(* Logix 5000 project; controller R400_500_XLS vendor 1 type 14 code 216 rev 31.11; software revision 31.01; part 29 of 32 *)
(* tags used below, declared in another part *)
   Abort1 : DINT;   // Not Used
   Alarm : SINT;   // Wait 3 seconds
   ClearIndex : DINT;
   Condenser : INT;
   CondenserHighFlow_1 : BOOL;   // Enables the condenser high flow valve
   CondenserHighFlow_2 : BOOL;   // Enables the condenser high flow valve
   CondenserLowFlow_1 : BOOL;   // Enables the condenser low flow valve
   CondenserLowFlow_2 : BOOL;   // Enables the condenser low flow valve
   CondenserTran : INT;
   CycleSequence : UDT_CYCLE_SEQUENCE;
   DrnSmp : DINT;
   DRYING : DINT;   // Drying id number
   F1rinse : DINT;   // Not Used
   F2rinse : DINT;   // Not Used
   F3rinse : DINT;   // Not Used
   FC06_ONS : DINT;
   FC06Tran1 : BOOL;   // Condition for the wash treatment to start
   FC07Tran1 : BOOL;   // Condition for the rinse treatment to start
   HeatSmp : DINT;
   iFindCRLFIndex : INT;   // Index Of CRLF in String
   iIndexClearMessageOverflowBuffer : INT;   // Message Overflow Buffer is sPrntArray(200-300)
   M : DINT[5];   // Memory Bits
   MinPressRecord : REAL;
   NeutralizationPhaseRequired : BOOL;
   OneShot : DINT[1];
   ONS_FC07 : SINT;
   print_Footer_template : STRING[7];   // Template for the cycle footer
   printTreatString : STRING[85];   // Treatment String
   rIn_WSH61 : REAL;
   Run : DINT;
   sCRLF : STRING;
   Service : DINT[2];   // Unused Service Mode Memory Bit
   sFll_Zero : STRING[20];
   sMessageToPrint : STRING;   // Message To Print
   sOut_WSH61 : STRING;
   sPrntArray : STRING[300];   // Printer String Array
   sResetPrinter : STRING;   // Clears Printer buffer jplv04f ASCII
   sSpaceCharacter : STRING;   // Space Character
   String : STRING[50];   // String
   SumpHeatingStopped : BOOL;   // Sump heating falling edge
   Tmr : TIMER[107];
   Trt_Drying : SINT;
   Trt_PrWsh : DINT;
   Trt_Rinse : DINT;   // Rinse steps
   Trt_Vapor_Exhaust : BOOL;   // Vapor exhaust fan is on
   Trt_Wsh : DINT;
   WSH56_StartHeating : BOOL;   // Start heating
   WSH56_StartPump : BOOL;   // Start pump signal
   WSH56_StartRecirculation : BOOL;   // Start the recirculation
   WSH_35 : BOOL;   // End of neutralization phase
   WshExcBuffer : UDT_WASH;
   AlarmTrigger : INT;   // Triggers the alarm screen if different of 0
   bCycleOrAbortInProcess : BOOL;
   bNewStringDetected : BOOL;
   DateFormat : SINT;   // 0: M-D-Y 1: D-M-Y 2: Y-M-D
   DateTime : DINT[7];
   ENABLE : BOOL;   // Enable bit
   EnaDisPrinter : BOOL;   // Screen 80 Enable/Disable Printer button
   PmpPres : REAL;
   PressureUnit : BOOL;   // Pressure Unit 0=PSIG 1=BAR
   printAlarm : STRING;
   printAlarmMsg : STRING[50];
   PrintChemCondValue : REAL;
   printEvent : STRING[5];
   PrintFrinseCondValue : REAL;
   PrintIndex : DINT;
   sDate : STRING;   // String current date
   sDateTime : STRING;   // String Date Time
   sNullCharacters : STRING;   // Empty String
   SPV_19 : BOOL;   // Screen 80 Enabled/Disabled Pump pressure monitoring
   sTime : STRING;   // String current time
   SumpTemp : REAL;   // Sump temperature in °C
   tStringCopyDebounce : TIMER;
   udtCSVDataLogBatchReport : UDT_CSVDataLog;
   Unit : Hrdwre;   // Unit Configuration
(* MainProgram, continued *)

ROUTINE WSH_56_TRT_WSH   (* ladder *)
// This module calls the routine to perform Wash treatments
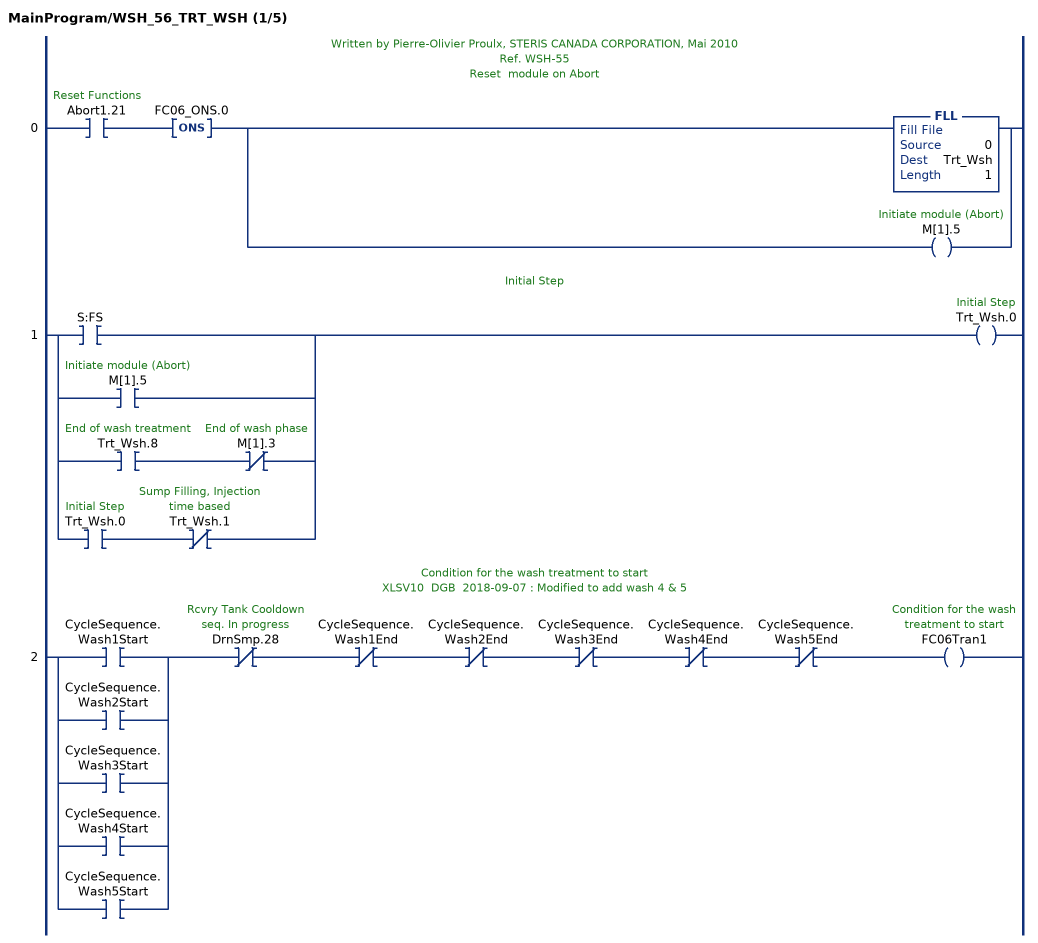
   // Written by Pierre-Olivier Proulx, STERIS CANADA CORPORATION, Mai 2010
   // Ref. WSH-55
   // Reset  module on Abort
   0: XIC(Abort1.21)ONS(FC06_ONS.0)[FLL(0,Trt_Wsh,1) ,OTE(M[1].5) ];
   // Initial Step
   1: [XIC(S:FS) ,XIC(M[1].5) ,XIC(Trt_Wsh.8) XIO(M[1].3) ,XIC(Trt_Wsh.0) XIO(Trt_Wsh.1) ]OTE(Trt_Wsh.0);
   // Condition for the wash treatment to start
   // XLSV10  DGB  2018-09-07 : Modified to add wash 4 & 5
   2: [XIC(CycleSequence.Wash1Start) ,XIC(CycleSequence.Wash2Start) ,XIC(CycleSequence.Wash3Start) ,XIC(CycleSequence.Wash4Start) ,XIC(CycleSequence.Wash5Start) ]XIO(DrnSmp.28)XIO(CycleSequence.Wash1End)XIO(CycleSequence.Wash2End)XIO(CycleSequence.Wash3End)XIO(CycleSequence.Wash4End)XIO(CycleSequence.Wash5End)OTE(FC06Tran1);
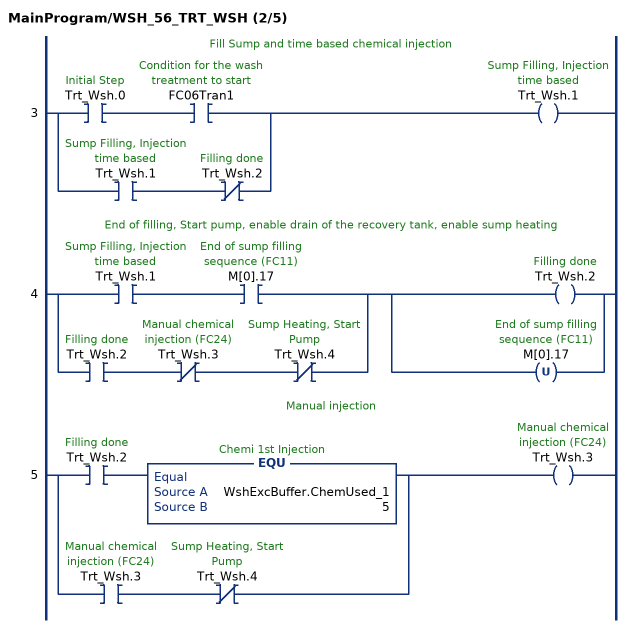
   // Fill Sump and time based chemical injection
   3: [XIC(Trt_Wsh.0) XIC(FC06Tran1) ,XIC(Trt_Wsh.1) XIO(Trt_Wsh.2) ]OTE(Trt_Wsh.1);
   // End of filling, Start pump, enable drain of the recovery tank, enable sump heating
   4: [XIC(Trt_Wsh.1) XIC(M[0].17) ,XIC(Trt_Wsh.2) XIO(Trt_Wsh.3) XIO(Trt_Wsh.4) ][OTE(Trt_Wsh.2) ,OTU(M[0].17) ];
   // Manual injection
   5: [XIC(Trt_Wsh.2) EQU(WshExcBuffer.ChemUsed_1,5) ,XIC(Trt_Wsh.3) XIO(Trt_Wsh.4) ]OTE(Trt_Wsh.3);
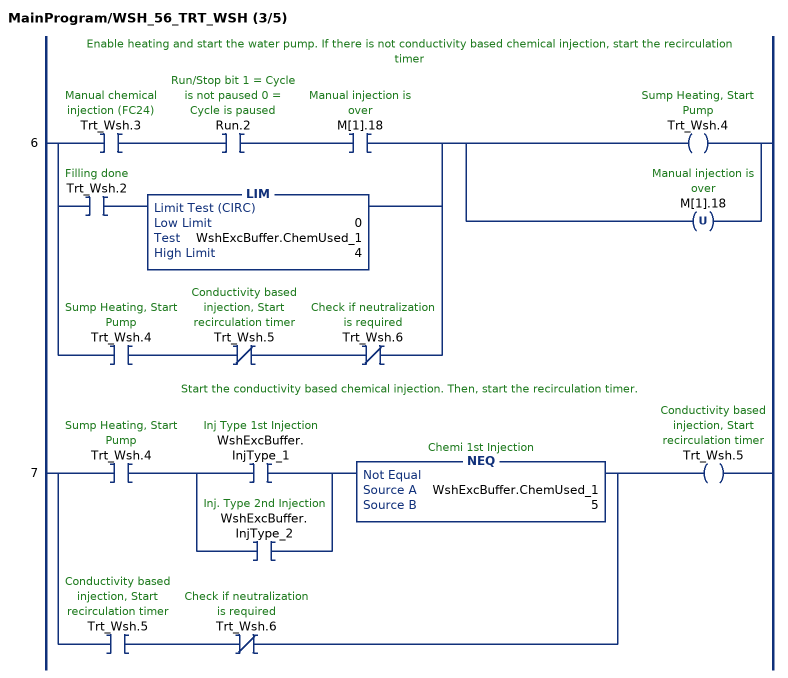
   // Enable heating and start the water pump. If there is not conductivity based chemical injection, start the recirculation timer
   6: [XIC(Trt_Wsh.3) XIC(Run.2) XIC(M[1].18) ,XIC(Trt_Wsh.2) LIM(0,WshExcBuffer.ChemUsed_1,4) ,XIC(Trt_Wsh.4) XIO(Trt_Wsh.5) XIO(Trt_Wsh.6) ][OTE(Trt_Wsh.4) ,OTU(M[1].18) ];
   // Start the conductivity based chemical injection. Then, start the recirculation timer.
   7: [XIC(Trt_Wsh.4) [XIC(WshExcBuffer.InjType_1) ,XIC(WshExcBuffer.InjType_2) ] NEQ(WshExcBuffer.ChemUsed_1,5) ,XIC(Trt_Wsh.5) XIO(Trt_Wsh.6) ]OTE(Trt_Wsh.5);
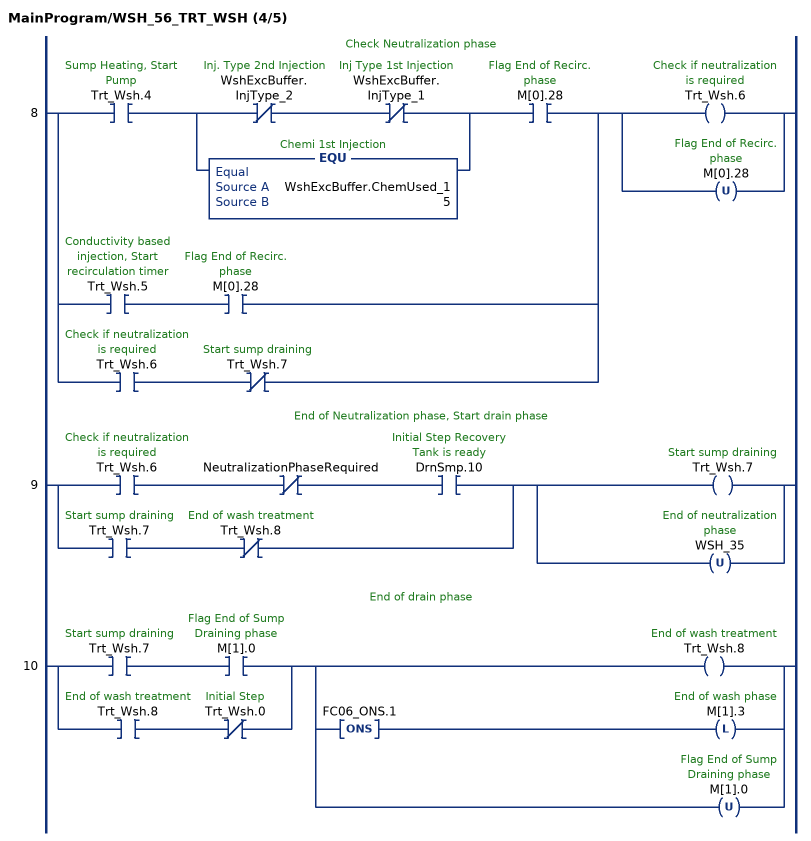
   // Check Neutralization phase
   8: [XIC(Trt_Wsh.4) [XIO(WshExcBuffer.InjType_2) XIO(WshExcBuffer.InjType_1) ,EQU(WshExcBuffer.ChemUsed_1,5) ] XIC(M[0].28) ,XIC(Trt_Wsh.5) XIC(M[0].28) ,XIC(Trt_Wsh.6) XIO(Trt_Wsh.7) ][OTE(Trt_Wsh.6) ,OTU(M[0].28) ];
   // End of Neutralization phase, Start drain phase
   9: [XIC(Trt_Wsh.6) XIO(NeutralizationPhaseRequired) XIC(DrnSmp.10) ,XIC(Trt_Wsh.7) XIO(Trt_Wsh.8) ][OTE(Trt_Wsh.7) ,OTU(WSH_35) ];
   // End of drain phase
   10: [XIC(Trt_Wsh.7) XIC(M[1].0) ,XIC(Trt_Wsh.8) XIO(Trt_Wsh.0) ][OTE(Trt_Wsh.8) ,ONS(FC06_ONS.1) OTL(M[1].3) ,OTU(M[1].0) ];
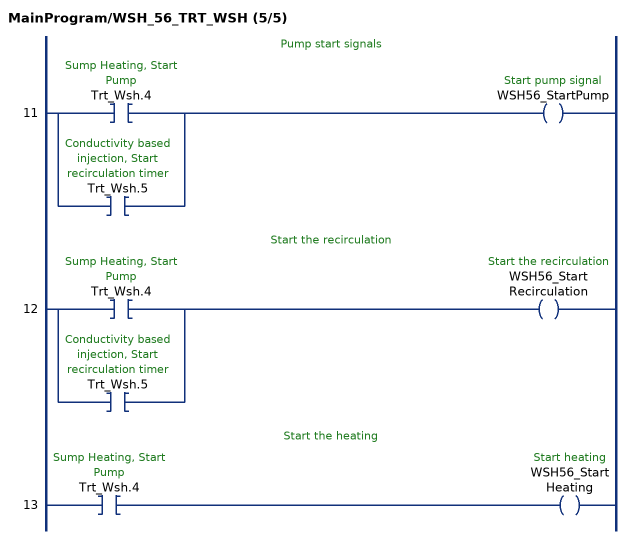
   // Pump start signals
   11: [XIC(Trt_Wsh.4) ,XIC(Trt_Wsh.5) ]OTE(WSH56_StartPump);
   // Start the recirculation
   12: [XIC(Trt_Wsh.4) ,XIC(Trt_Wsh.5) ]OTE(WSH56_StartRecirculation);
   // Start the heating
   13: XIC(Trt_Wsh.4)OTE(WSH56_StartHeating);
END_ROUTINE

ROUTINE WSH_57_TRT_RINSE   (* ladder *)
// This routine performs a rinse treatment.
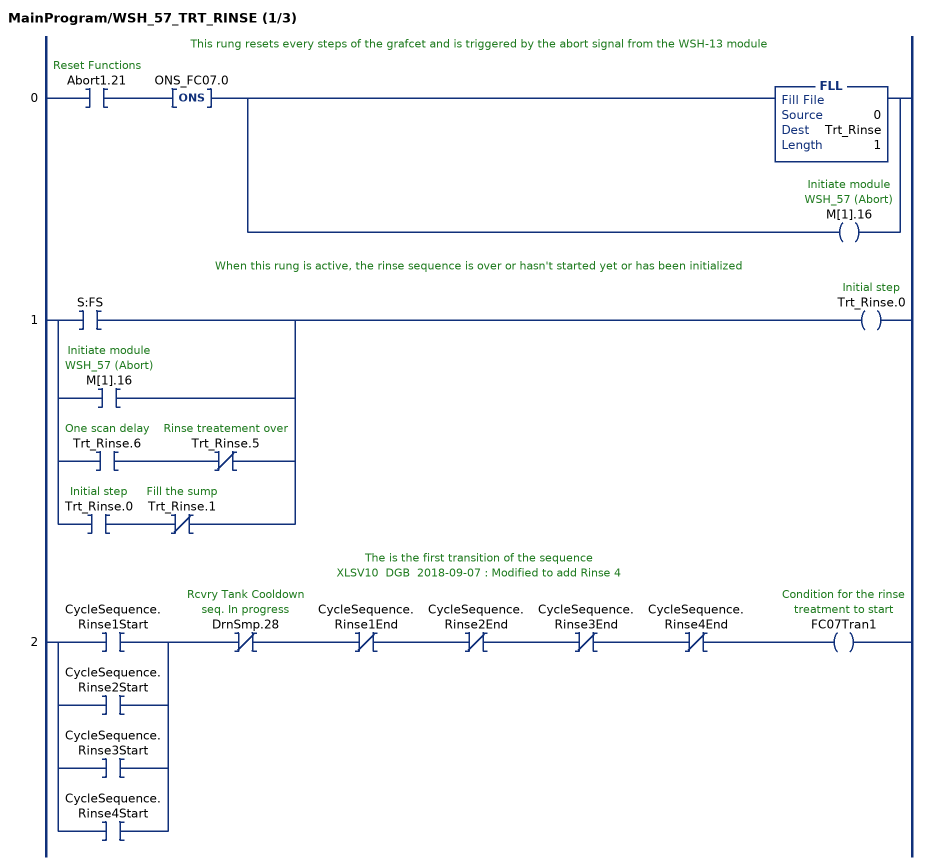
   // This rung resets every steps of the grafcet and is triggered by the abort signal from the WSH-13 module
   0: XIC(Abort1.21)ONS(ONS_FC07.0)[FLL(0,Trt_Rinse,1) ,OTE(M[1].16) ];
   // When this rung is active, the rinse sequence is over or hasn't started yet or has been initialized
   1: [XIC(S:FS) ,XIC(M[1].16) ,XIC(Trt_Rinse.6) XIO(Trt_Rinse.5) ,XIC(Trt_Rinse.0) XIO(Trt_Rinse.1) ]OTE(Trt_Rinse.0);
   // The is the first transition of the sequence
   // XLSV10  DGB  2018-09-07 : Modified to add Rinse 4
   2: [XIC(CycleSequence.Rinse1Start) ,XIC(CycleSequence.Rinse2Start) ,XIC(CycleSequence.Rinse3Start) ,XIC(CycleSequence.Rinse4Start) ]XIO(DrnSmp.28)XIO(CycleSequence.Rinse1End)XIO(CycleSequence.Rinse2End)XIO(CycleSequence.Rinse3End)XIO(CycleSequence.Rinse4End)OTE(FC07Tran1);
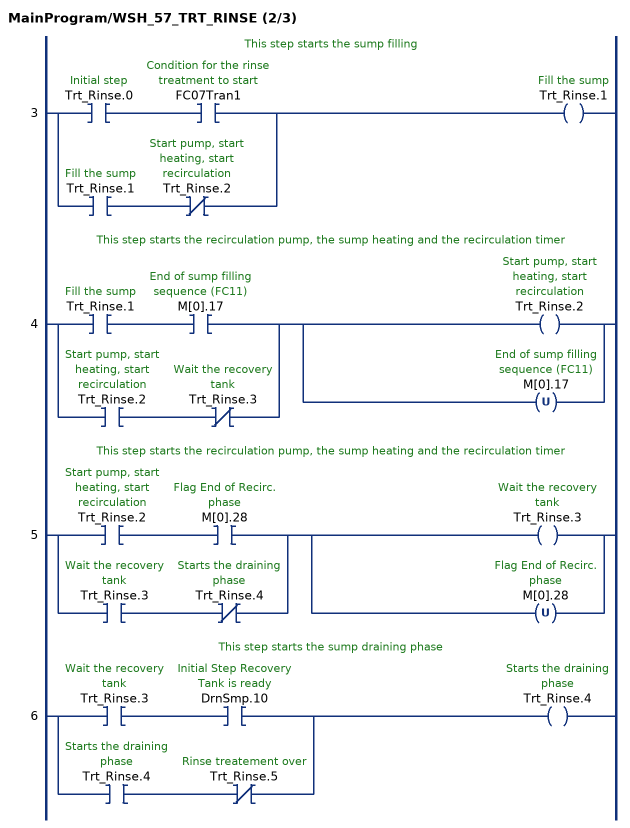
   // This step starts the sump filling
   3: [XIC(Trt_Rinse.0) XIC(FC07Tran1) ,XIC(Trt_Rinse.1) XIO(Trt_Rinse.2) ]OTE(Trt_Rinse.1);
   // This step starts the recirculation pump, the sump heating and the recirculation timer
   4: [XIC(Trt_Rinse.1) XIC(M[0].17) ,XIC(Trt_Rinse.2) XIO(Trt_Rinse.3) ][OTE(Trt_Rinse.2) ,OTU(M[0].17) ];
   // This step starts the recirculation pump, the sump heating and the recirculation timer
   5: [XIC(Trt_Rinse.2) XIC(M[0].28) ,XIC(Trt_Rinse.3) XIO(Trt_Rinse.4) ][OTE(Trt_Rinse.3) ,OTU(M[0].28) ];
   // This step starts the sump draining phase
   6: [XIC(Trt_Rinse.3) XIC(DrnSmp.10) ,XIC(Trt_Rinse.4) XIO(Trt_Rinse.5) ]OTE(Trt_Rinse.4);
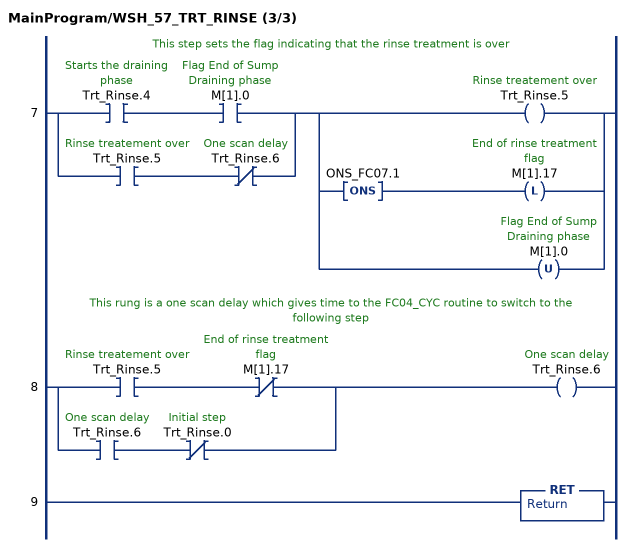
   // This step sets the flag indicating that the rinse treatment is over
   7: [XIC(Trt_Rinse.4) XIC(M[1].0) ,XIC(Trt_Rinse.5) XIO(Trt_Rinse.6) ][OTE(Trt_Rinse.5) ,ONS(ONS_FC07.1) OTL(M[1].17) ,OTU(M[1].0) ];
   // This rung is a one scan delay which gives time to the FC04_CYC routine to switch to the following step
   8: [XIC(Trt_Rinse.5) XIO(M[1].17) ,XIC(Trt_Rinse.6) XIO(Trt_Rinse.0) ]OTE(Trt_Rinse.6);
   9: RET();
END_ROUTINE

ROUTINE WSH_59_CONDENSER_WET   (* ladder *)
// This routine manages the condenser operation
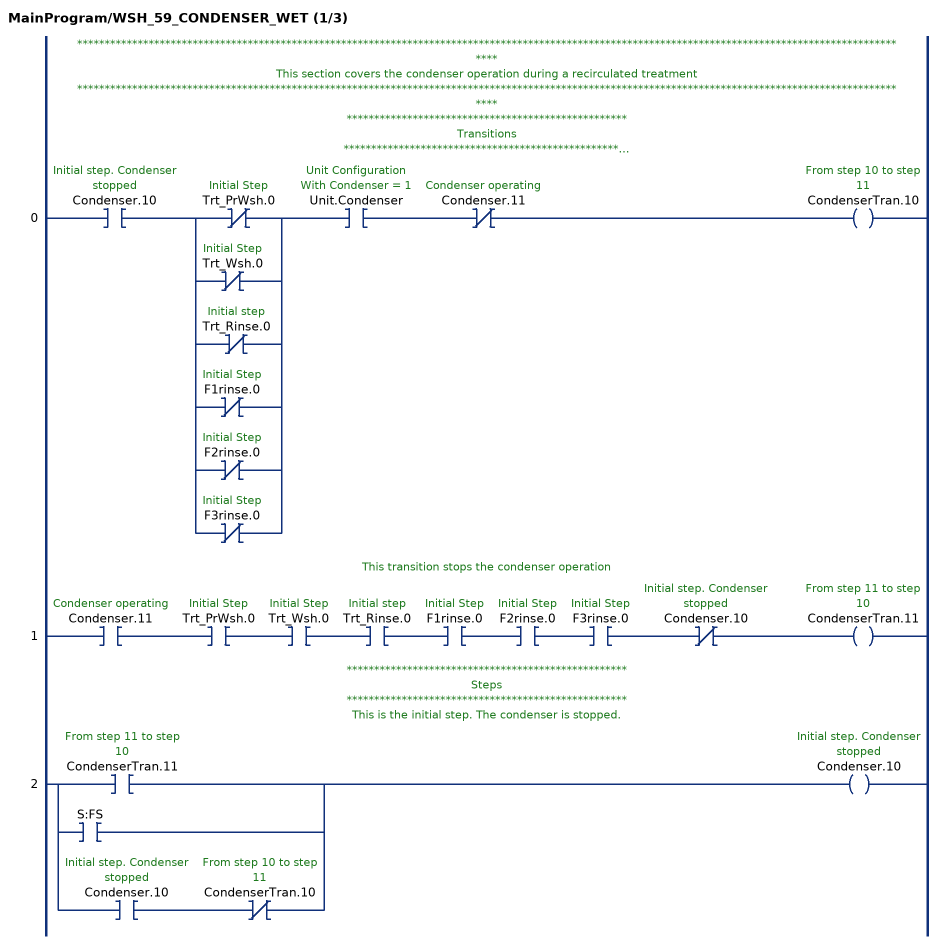
   // *********************************************************************************************************************************************************
   // This section covers the condenser operation during a recirculated treatment
   // *********************************************************************************************************************************************************
   // ***************************************************
   // Transitions
   // ***************************************************
   // This condition triggers the condenser operation
   0: XIC(Condenser.10)[XIO(Trt_PrWsh.0) ,XIO(Trt_Wsh.0) ,XIO(Trt_Rinse.0) ,XIO(F1rinse.0) ,XIO(F2rinse.0) ,XIO(F3rinse.0) ]XIC(Unit.Condenser)XIO(Condenser.11)OTE(CondenserTran.10);
   // This transition stops the condenser operation
   1: XIC(Condenser.11)XIC(Trt_PrWsh.0)XIC(Trt_Wsh.0)XIC(Trt_Rinse.0)XIC(F1rinse.0)XIC(F2rinse.0)XIC(F3rinse.0)XIO(Condenser.10)OTE(CondenserTran.11);
   // ***************************************************
   // Steps
   // ***************************************************
   // This is the initial step. The condenser is stopped.
   2: [XIC(CondenserTran.11) ,XIC(S:FS) ,XIC(Condenser.10) XIO(CondenserTran.10) ]OTE(Condenser.10);
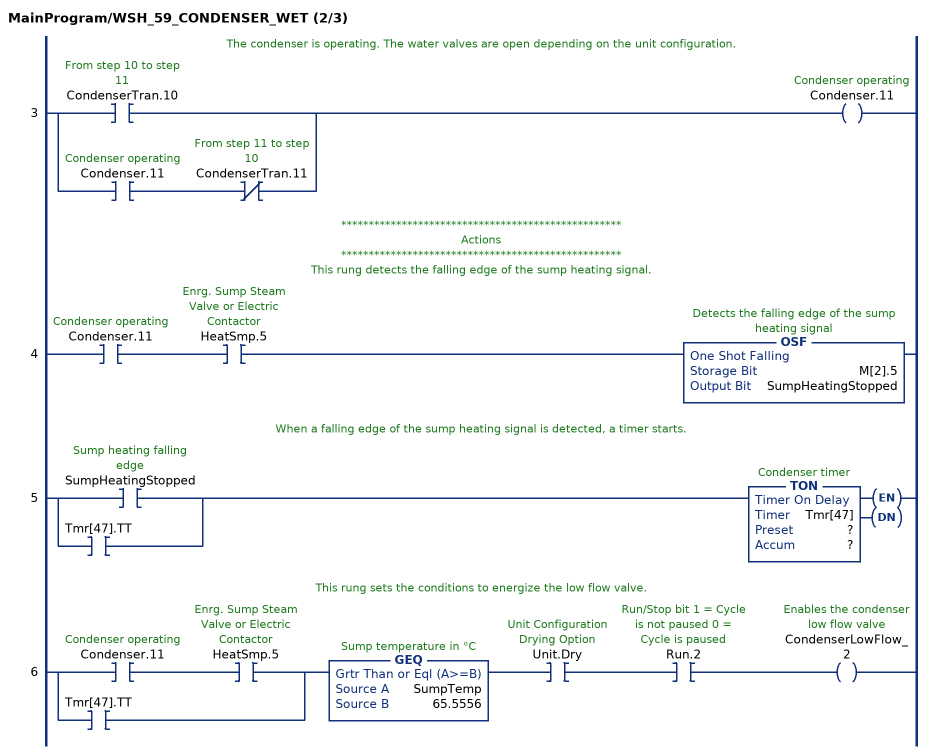
   // The condenser is operating. The water valves are open depending on the unit configuration.
   3: [XIC(CondenserTran.10) ,XIC(Condenser.11) XIO(CondenserTran.11) ]OTE(Condenser.11);
   // ***************************************************
   // Actions
   // ***************************************************
   // This rung detects the falling edge of the sump heating signal.
   4: XIC(Condenser.11)XIC(HeatSmp.5)OSF(M[2].5,SumpHeatingStopped);
   // When a falling edge of the sump heating signal is detected, a timer starts.
   5: [XIC(SumpHeatingStopped) ,XIC(Tmr[47].TT) ]TON(Tmr[47],?,?);
   // This rung sets the conditions to energize the low flow valve.
   6: [XIC(Condenser.11) XIC(HeatSmp.5) ,XIC(Tmr[47].TT) ]GEQ(SumpTemp,65.5556)XIC(Unit.Dry)XIC(Run.2)OTE(CondenserLowFlow_2);
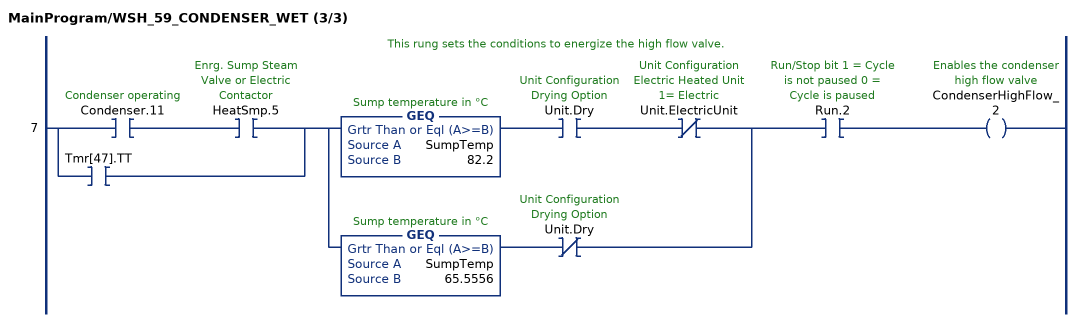
   // This rung sets the conditions to energize the high flow valve.
   7: [XIC(Condenser.11) XIC(HeatSmp.5) ,XIC(Tmr[47].TT) ][GEQ(SumpTemp,82.2) XIC(Unit.Dry) XIO(Unit.ElectricUnit) ,GEQ(SumpTemp,65.5556) XIO(Unit.Dry) ]XIC(Run.2)OTE(CondenserHighFlow_2);
END_ROUTINE

ROUTINE WSH_60_CONDENSER_DRY_VENT   (* ladder *)
// This routine manages the condenser operation
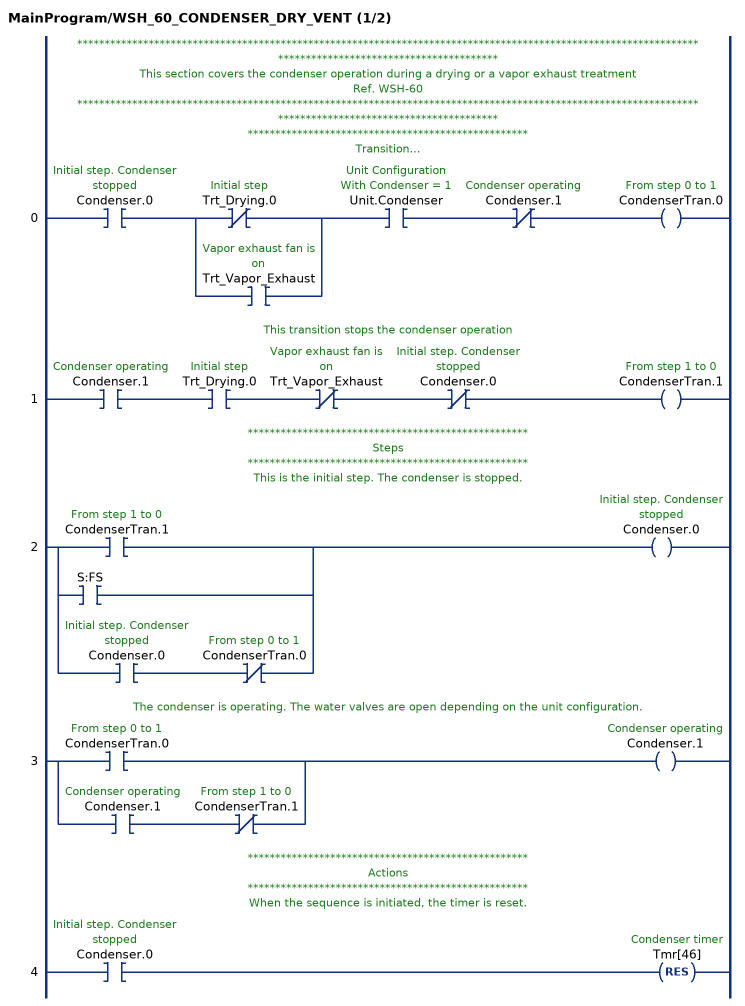
   // *********************************************************************************************************************************************************
   // This section covers the condenser operation during a drying or a vapor exhaust treatment
   // Ref. WSH-60
   // *********************************************************************************************************************************************************
   // ***************************************************
   // Transitions
   // ***************************************************
   // This condition triggers the condenser operation
   0: XIC(Condenser.0)[XIO(Trt_Drying.0) ,XIC(Trt_Vapor_Exhaust) ]XIC(Unit.Condenser)XIO(Condenser.1)OTE(CondenserTran.0);
   // This transition stops the condenser operation
   1: XIC(Condenser.1)XIC(Trt_Drying.0)XIO(Trt_Vapor_Exhaust)XIO(Condenser.0)OTE(CondenserTran.1);
   // ***************************************************
   // Steps
   // ***************************************************
   // This is the initial step. The condenser is stopped.
   2: [XIC(CondenserTran.1) ,XIC(S:FS) ,XIC(Condenser.0) XIO(CondenserTran.0) ]OTE(Condenser.0);
   // The condenser is operating. The water valves are open depending on the unit configuration.
   3: [XIC(CondenserTran.0) ,XIC(Condenser.1) XIO(CondenserTran.1) ]OTE(Condenser.1);
   // ***************************************************
   // Actions
   // ***************************************************
   // When the sequence is initiated, the timer is reset.
   4: XIC(Condenser.0)RES(Tmr[46]);
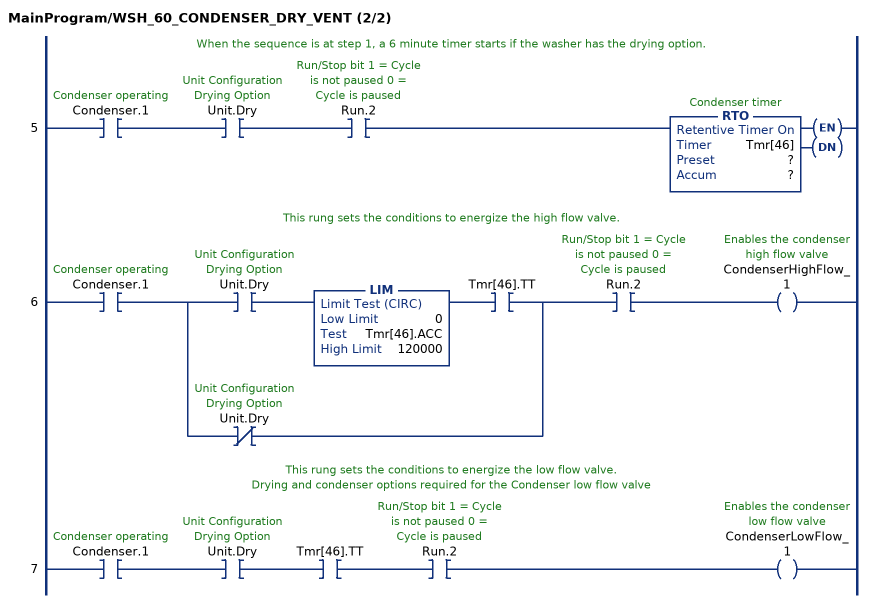
   // When the sequence is at step 1, a 6 minute timer starts if the washer has the drying option.
   5: XIC(Condenser.1)XIC(Unit.Dry)XIC(Run.2)RTO(Tmr[46],?,?);
   // This rung sets the conditions to energize the high flow valve.
   6: XIC(Condenser.1)[XIC(Unit.Dry) LIM(0,Tmr[46].ACC,120000) XIC(Tmr[46].TT) ,XIO(Unit.Dry) ]XIC(Run.2)OTE(CondenserHighFlow_1);
   // This rung sets the conditions to energize the low flow valve.
   // Drying and condenser options required for the Condenser low flow valve
   7: XIC(Condenser.1)XIC(Unit.Dry)XIC(Tmr[46].TT)XIC(Run.2)OTE(CondenserLowFlow_1);
END_ROUTINE

ROUTINE WSH_61_PRINT_STRING_ELEMENT   (* ladder *)
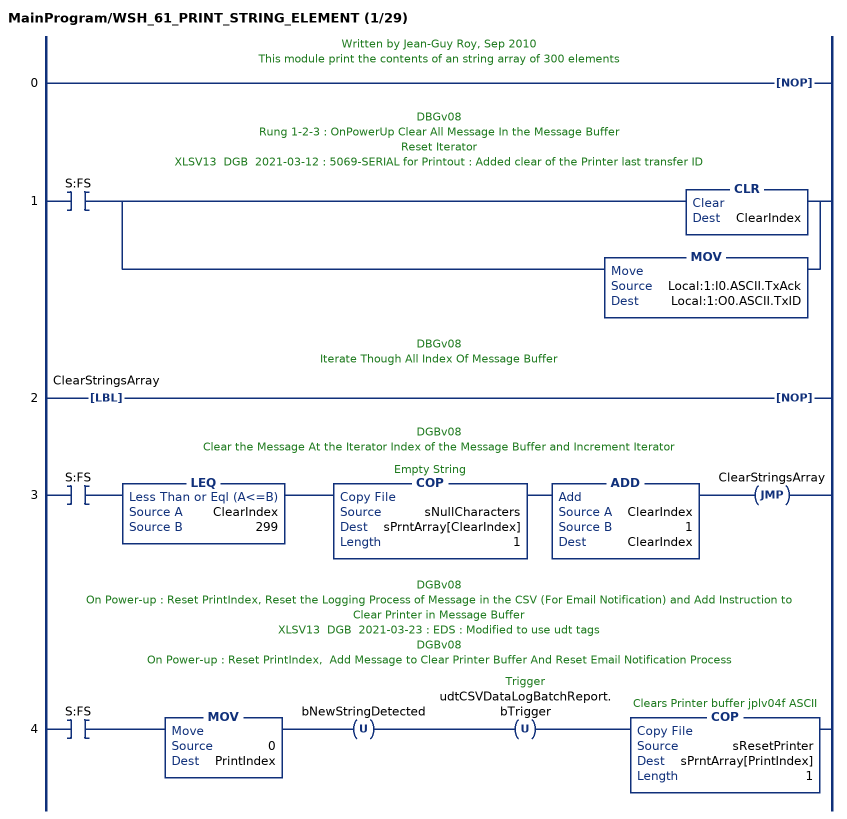
   // Written by Jean-Guy Roy, Sep 2010
   // This module print the contents of an string array of 300 elements
   0: NOP();
   // DBGv08
   // Rung 1-2-3 : OnPowerUp Clear All Message In the Message Buffer
   // Reset Iterator
   // XLSV13  DGB  2021-03-12 : 5069-SERIAL for Printout : Added clear of the Printer last transfer ID
   1: XIC(S:FS)[CLR(ClearIndex) ,MOV(Local:1:I0.ASCII.TxAck,Local:1:O0.ASCII.TxID) ];
   // DBGv08
   // Iterate Though All Index Of Message Buffer
   2: LBL(ClearStringsArray)NOP();
   // DGBv08
   // Clear the Message At the Iterator Index of the Message Buffer and Increment Iterator
   3: XIC(S:FS)LEQ(ClearIndex,299)COP(sNullCharacters,sPrntArray[ClearIndex],1)ADD(ClearIndex,1,ClearIndex)JMP(ClearStringsArray);
   // DGBv08
   // On Power-up : Reset PrintIndex, Reset the Logging Process of Message in the CSV (For Email Notification) and Add Instruction to Clear Printer in Message Buffer
   // XLSV13  DGB  2021-03-23 : EDS : Modified to use udt tags
   // DGBv08
   // On Power-up : Reset PrintIndex,  Add Message to Clear Printer Buffer And Reset Email Notification Process
   4: XIC(S:FS)MOV(0,PrintIndex)OTU(bNewStringDetected)OTU(udtCSVDataLogBatchReport.bTrigger)COP(sResetPrinter,sPrntArray[PrintIndex],1);
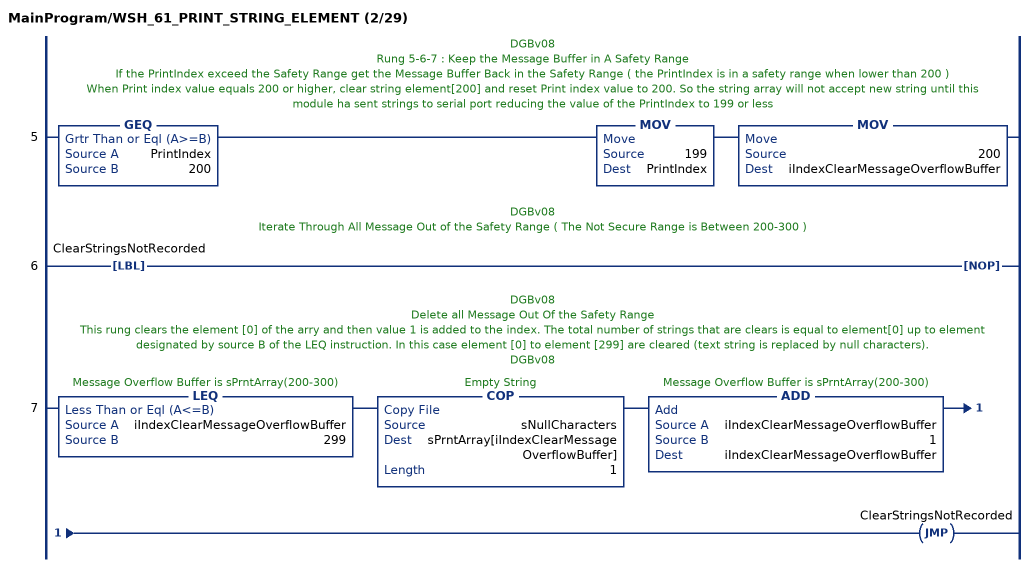
   // DGBv08
   // Rung 5-6-7 : Keep the Message Buffer in A Safety Range
   // If the PrintIndex exceed the Safety Range get the Message Buffer Back in the Safety Range ( the PrintIndex is in a safety range when lower than 200 )
   // When Print index value equals 200 or higher, clear string element[200] and reset Print index value to 200. So the string array will not accept new string until this module ha sent strings to serial port reducing the value of the PrintIndex to 199 or less
   5: GEQ(PrintIndex,200)MOV(199,PrintIndex)MOV(200,iIndexClearMessageOverflowBuffer);
   // DGBv08
   // Iterate Through All Message Out of the Safety Range ( The Not Secure Range is Between 200-300 )
   6: LBL(ClearStringsNotRecorded)NOP();
   // DGBv08
   // Delete all Message Out Of the Safety Range
   // This rung clears the element [0] of the arry and then value 1 is added to the index. The total number of strings that are clears is equal to element[0] up to element designated by source B of the LEQ instruction. In this case element [0] to element [299] are cleared (text string is replaced by null characters).
   // DGBv08
   7: LEQ(iIndexClearMessageOverflowBuffer,299)COP(sNullCharacters,sPrntArray[iIndexClearMessageOverflowBuffer],1)ADD(iIndexClearMessageOverflowBuffer,1,iIndexClearMessageOverflowBuffer)JMP(ClearStringsNotRecorded);
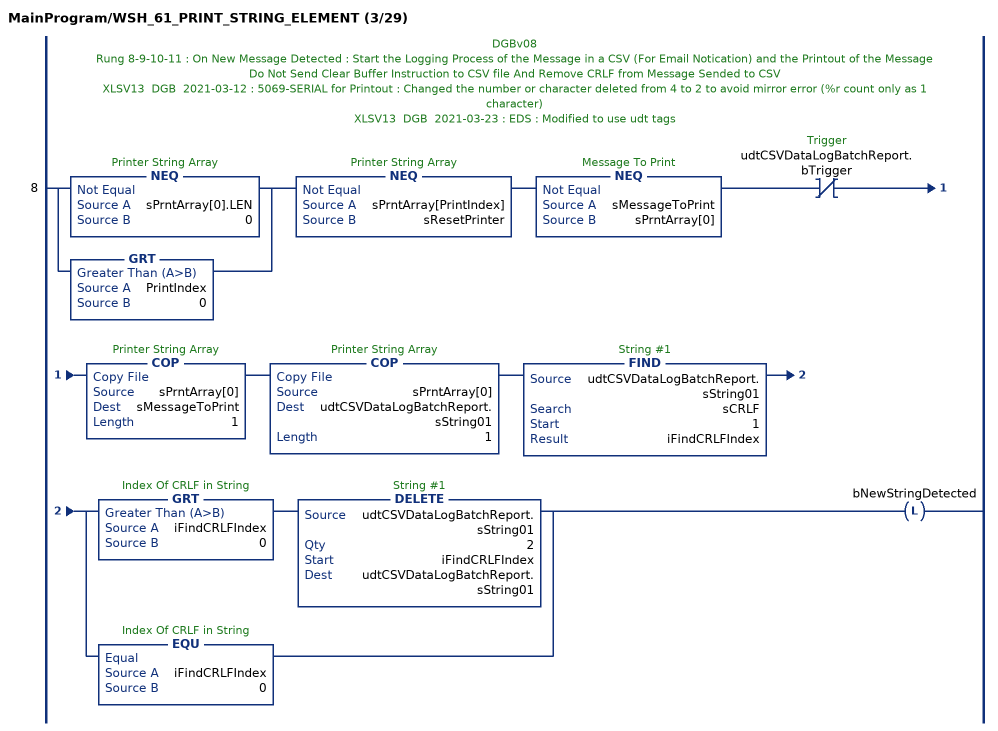
   // DGBv08
   // Rung 8-9-10-11 : On New Message Detected : Start the Logging Process of the Message in a CSV (For Email Notication) and the Printout of the Message
   // Do Not Send Clear Buffer Instruction to CSV file And Remove CRLF from Message Sended to CSV
   // XLSV13  DGB  2021-03-12 : 5069-SERIAL for Printout : Changed the number or character deleted from 4 to 2 to avoid mirror error (%r count only as 1 character)
   // XLSV13  DGB  2021-03-23 : EDS : Modified to use udt tags
   8: [NEQ(sPrntArray[0].LEN,0) ,GRT(PrintIndex,0) ]NEQ(sPrntArray[PrintIndex],sResetPrinter)NEQ(sMessageToPrint,sPrntArray[0])XIO(udtCSVDataLogBatchReport.bTrigger)COP(sPrntArray[0],sMessageToPrint,1)COP(sPrntArray[0],udtCSVDataLogBatchReport.sString01,1)FIND(udtCSVDataLogBatchReport.sString01,sCRLF,1,iFindCRLFIndex)[GRT(iFindCRLFIndex,0) DELETE(udtCSVDataLogBatchReport.sString01,2,iFindCRLFIndex,udtCSVDataLogBatchReport.sString01) ,EQU(iFindCRLFIndex,0) ]OTL(bNewStringDetected);
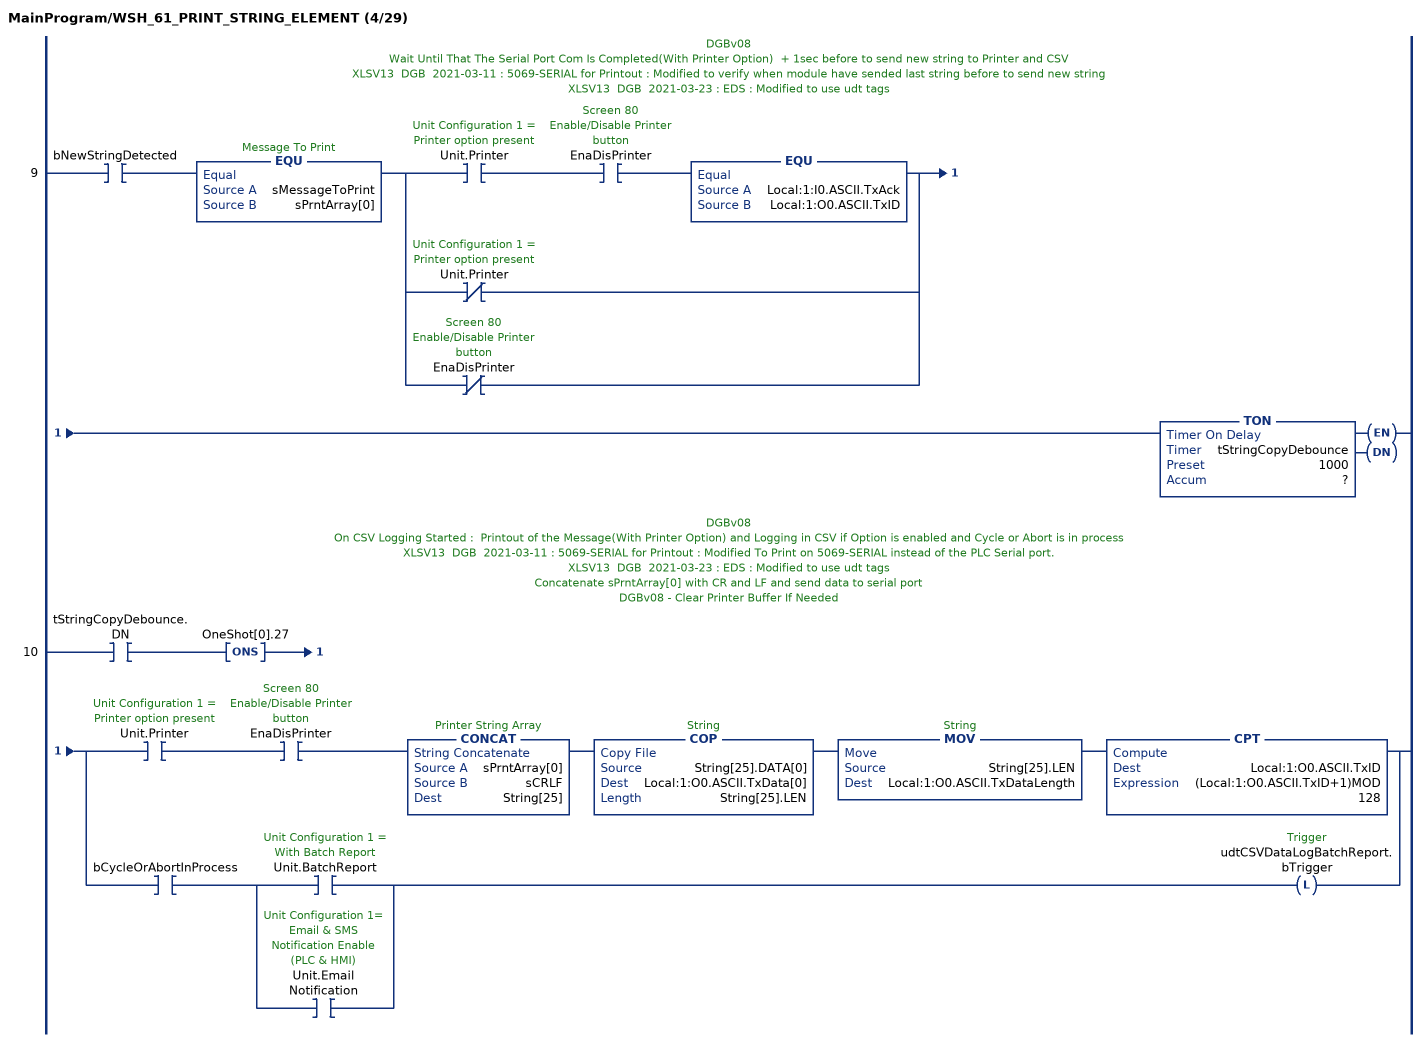
   // DGBv08
   // Wait Until That The Serial Port Com Is Completed(With Printer Option)  + 1sec before to send new string to Printer and CSV
   // XLSV13  DGB  2021-03-11 : 5069-SERIAL for Printout : Modified to verify when module have sended last string before to send new string
   // XLSV13  DGB  2021-03-23 : EDS : Modified to use udt tags
   9: XIC(bNewStringDetected)EQU(sMessageToPrint,sPrntArray[0])[XIC(Unit.Printer) XIC(EnaDisPrinter) EQU(Local:1:I0.ASCII.TxAck,Local:1:O0.ASCII.TxID) ,XIO(Unit.Printer) ,XIO(EnaDisPrinter) ]TON(tStringCopyDebounce,?,?);
   // DGBv08
   // On CSV Logging Started :  Printout of the Message(With Printer Option) and Logging in CSV if Option is enabled and Cycle or Abort is in process
   // XLSV13  DGB  2021-03-11 : 5069-SERIAL for Printout : Modified To Print on 5069-SERIAL instead of the PLC Serial port.
   // XLSV13  DGB  2021-03-23 : EDS : Modified to use udt tags
   // Concatenate sPrntArray[0] with CR and LF and send data to serial port
   // DGBv08 - Clear Printer Buffer If Needed
   10: XIC(tStringCopyDebounce.DN)ONS(OneShot[0].27)[XIC(Unit.Printer) XIC(EnaDisPrinter) CONCAT(sPrntArray[0],sCRLF,String[25]) COP(String[25].DATA[0],Local:1:O0.ASCII.TxData[0],String[25].LEN) MOV(String[25].LEN,Local:1:O0.ASCII.TxDataLength) CPT(Local:1:O0.ASCII.TxID,(Local:1:O0.ASCII.TxID+1)MOD 128) ,XIC(bCycleOrAbortInProcess) [XIC(Unit.BatchReport) ,XIC(Unit.EmailNotification) ] OTL(udtCSVDataLogBatchReport.bTrigger) ];
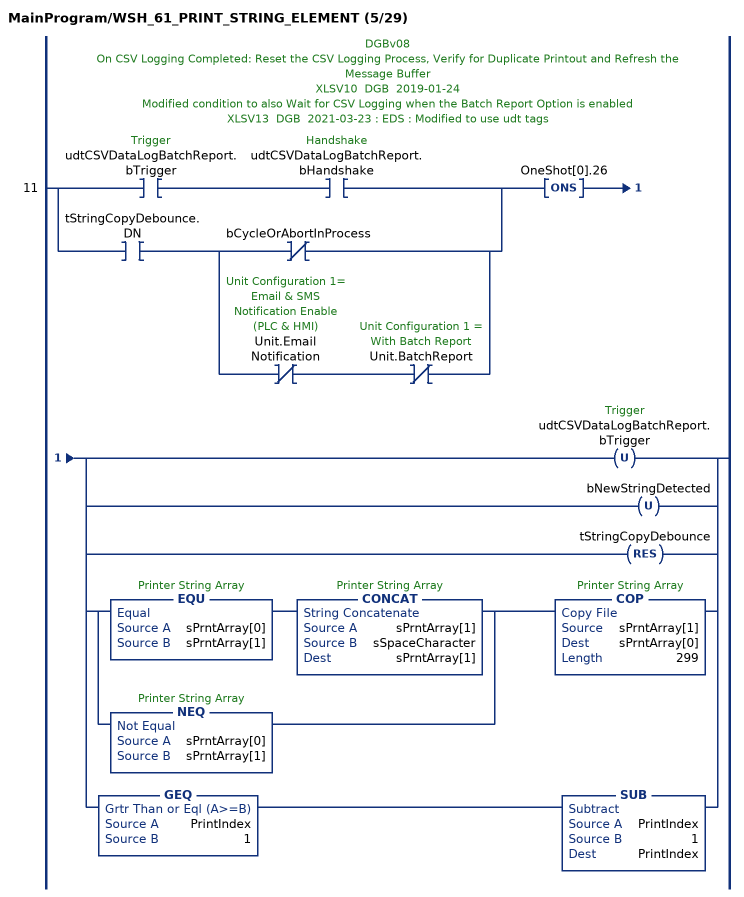
   // DGBv08
   // On CSV Logging Completed: Reset the CSV Logging Process, Verify for Duplicate Printout and Refresh the Message Buffer
   // XLSV10  DGB  2019-01-24
   // Modified condition to also Wait for CSV Logging when the Batch Report Option is enabled
   // XLSV13  DGB  2021-03-23 : EDS : Modified to use udt tags
   11: [XIC(udtCSVDataLogBatchReport.bTrigger) XIC(udtCSVDataLogBatchReport.bHandshake) ,XIC(tStringCopyDebounce.DN) [XIO(bCycleOrAbortInProcess) ,XIO(Unit.EmailNotification) XIO(Unit.BatchReport) ] ]ONS(OneShot[0].26)[OTU(udtCSVDataLogBatchReport.bTrigger) ,OTU(bNewStringDetected) ,RES(tStringCopyDebounce) ,[EQU(sPrntArray[0],sPrntArray[1]) CONCAT(sPrntArray[1],sSpaceCharacter,sPrntArray[1]) ,NEQ(sPrntArray[0],sPrntArray[1]) ] COP(sPrntArray[1],sPrntArray[0],299) ,GEQ(PrintIndex,1) SUB(PrintIndex,1,PrintIndex) ];
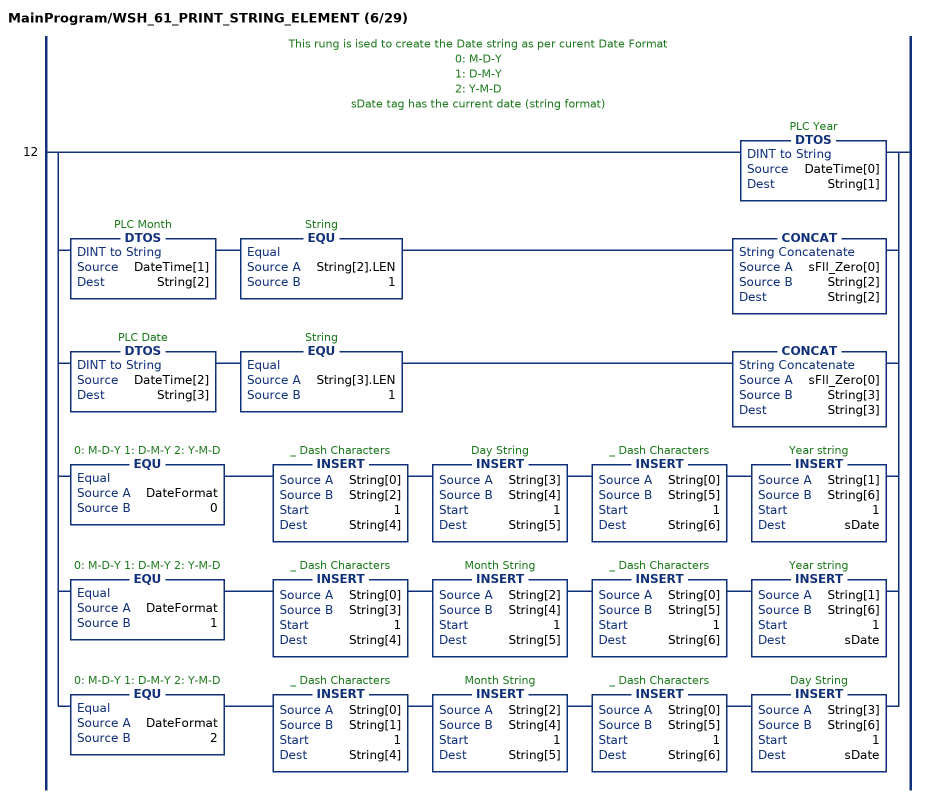
   // This rung is ised to create the Date string as per curent Date Format
   // 0: M-D-Y
   // 1: D-M-Y
   // 2: Y-M-D
   // sDate tag has the current date (string format)
   12: [DTOS(DateTime[0],String[1]) ,DTOS(DateTime[1],String[2]) EQU(String[2].LEN,1) CONCAT(sFll_Zero[0],String[2],String[2]) ,DTOS(DateTime[2],String[3]) EQU(String[3].LEN,1) CONCAT(sFll_Zero[0],String[3],String[3]) ,EQU(DateFormat,0) INSERT(String[0],String[2],1,String[4]) INSERT(String[3],String[4],1,String[5]) INSERT(String[0],String[5],1,String[6]) INSERT(String[1],String[6],1,sDate) ,EQU(DateFormat,1) INSERT(String[0],String[3],1,String[4]) INSERT(String[2],String[4],1,String[5]) INSERT(String[0],String[5],1,String[6]) INSERT(String[1],String[6],1,sDate) ,EQU(DateFormat,2) INSERT(String[0],String[1],1,String[4]) INSERT(String[2],String[4],1,String[5]) INSERT(String[0],String[5],1,String[6]) INSERT(String[3],String[6],1,sDate) ];
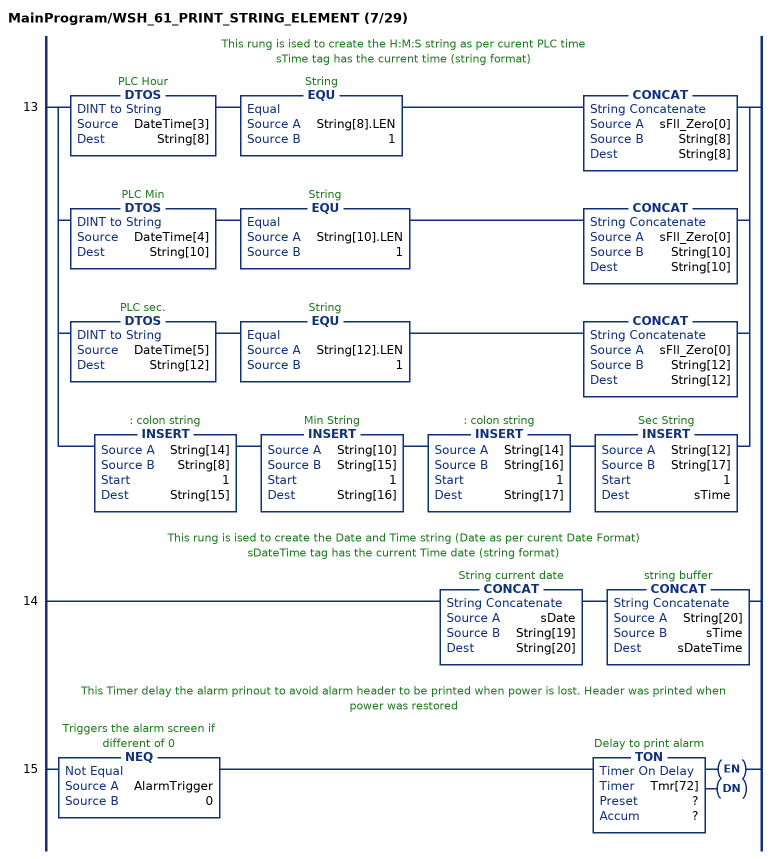
   // This rung is ised to create the H:M:S string as per curent PLC time
   // sTime tag has the current time (string format)
   13: [DTOS(DateTime[3],String[8]) EQU(String[8].LEN,1) CONCAT(sFll_Zero[0],String[8],String[8]) ,DTOS(DateTime[4],String[10]) EQU(String[10].LEN,1) CONCAT(sFll_Zero[0],String[10],String[10]) ,DTOS(DateTime[5],String[12]) EQU(String[12].LEN,1) CONCAT(sFll_Zero[0],String[12],String[12]) ,INSERT(String[14],String[8],1,String[15]) INSERT(String[10],String[15],1,String[16]) INSERT(String[14],String[16],1,String[17]) INSERT(String[12],String[17],1,sTime) ];
   // This rung is ised to create the Date and Time string (Date as per curent Date Format)
   // sDateTime tag has the current Time date (string format)
   14: CONCAT(sDate,String[19],String[20])CONCAT(String[20],sTime,sDateTime);
   // This Timer delay the alarm prinout to avoid alarm header to be printed when power is lost. Header was printed when power was restored
   15: NEQ(AlarmTrigger,0)TON(Tmr[72],?,?);
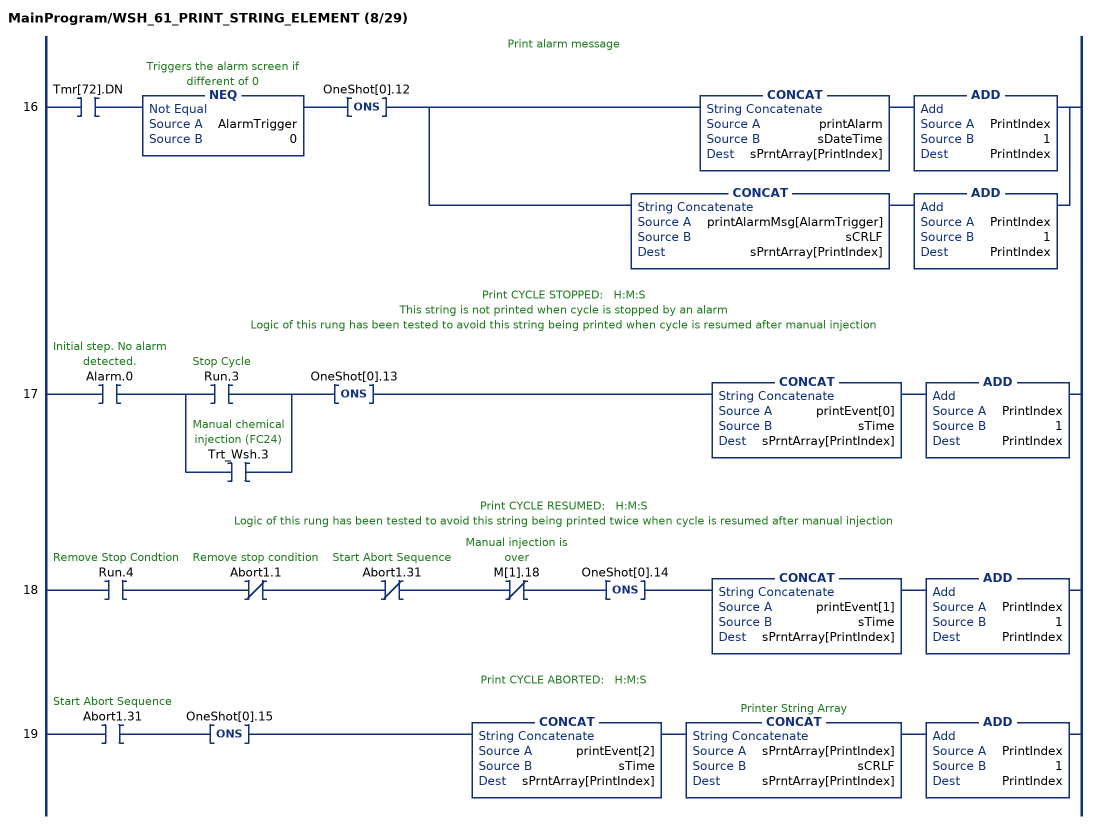
   // Print alarm message
   16: XIC(Tmr[72].DN)NEQ(AlarmTrigger,0)ONS(OneShot[0].12)[CONCAT(printAlarm,sDateTime,sPrntArray[PrintIndex]) ADD(PrintIndex,1,PrintIndex) ,CONCAT(printAlarmMsg[AlarmTrigger],sCRLF,sPrntArray[PrintIndex]) ADD(PrintIndex,1,PrintIndex) ];
   // Print CYCLE STOPPED:   H:M:S
   // This string is not printed when cycle is stopped by an alarm
   // Logic of this rung has been tested to avoid this string being printed when cycle is resumed after manual injection
   17: XIC(Alarm.0)[XIC(Run.3) ,XIC(Trt_Wsh.3) ]ONS(OneShot[0].13)CONCAT(printEvent[0],sTime,sPrntArray[PrintIndex])ADD(PrintIndex,1,PrintIndex);
   // Print CYCLE RESUMED:   H:M:S
   // Logic of this rung has been tested to avoid this string being printed twice when cycle is resumed after manual injection
   18: XIC(Run.4)XIO(Abort1.1)XIO(Abort1.31)XIO(M[1].18)ONS(OneShot[0].14)CONCAT(printEvent[1],sTime,sPrntArray[PrintIndex])ADD(PrintIndex,1,PrintIndex);
   // Print CYCLE ABORTED:   H:M:S
   19: XIC(Abort1.31)ONS(OneShot[0].15)CONCAT(printEvent[2],sTime,sPrntArray[PrintIndex])CONCAT(sPrntArray[PrintIndex],sCRLF,sPrntArray[PrintIndex])ADD(PrintIndex,1,PrintIndex);
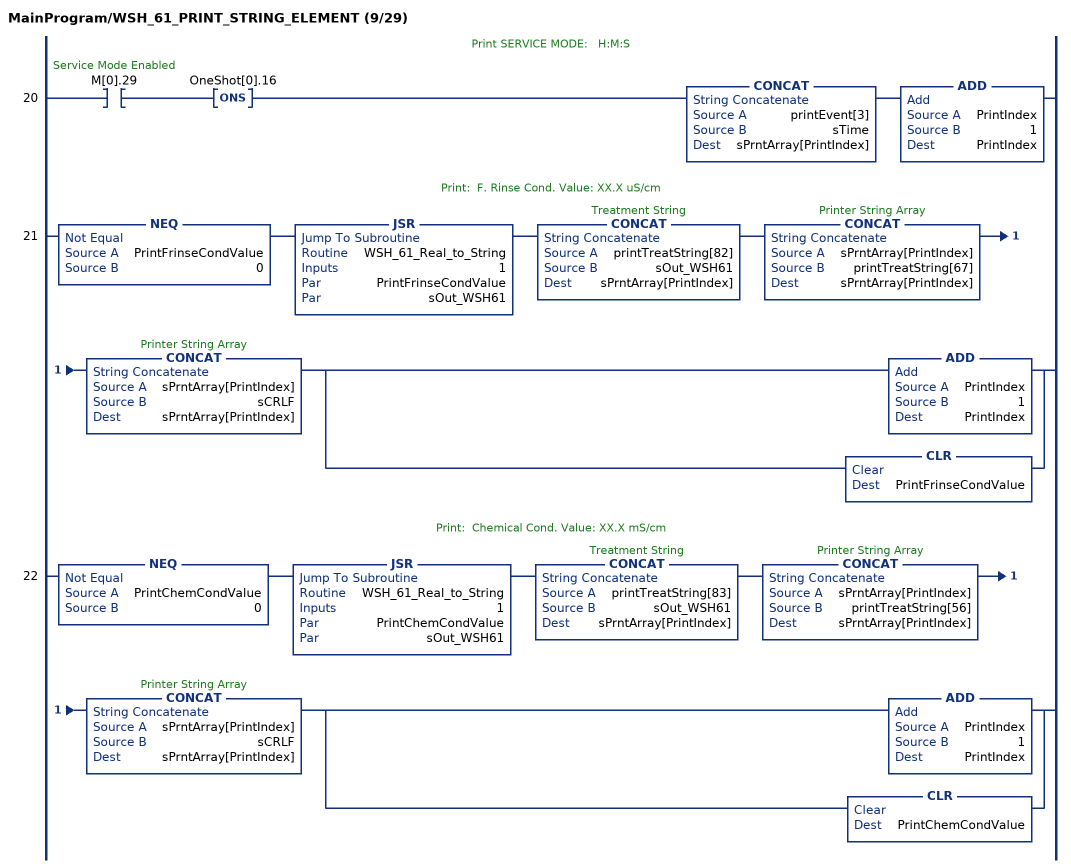
   // Print SERVICE MODE:   H:M:S
   20: XIC(M[0].29)ONS(OneShot[0].16)CONCAT(printEvent[3],sTime,sPrntArray[PrintIndex])ADD(PrintIndex,1,PrintIndex);
   // Print:  F. Rinse Cond. Value: XX.X uS/cm
   21: NEQ(PrintFrinseCondValue,0)JSR(WSH_61_Real_to_String,1,PrintFrinseCondValue,sOut_WSH61)CONCAT(printTreatString[82],sOut_WSH61,sPrntArray[PrintIndex])CONCAT(sPrntArray[PrintIndex],printTreatString[67],sPrntArray[PrintIndex])CONCAT(sPrntArray[PrintIndex],sCRLF,sPrntArray[PrintIndex])[ADD(PrintIndex,1,PrintIndex) ,CLR(PrintFrinseCondValue) ];
   // Print:  Chemical Cond. Value: XX.X mS/cm
   22: NEQ(PrintChemCondValue,0)JSR(WSH_61_Real_to_String,1,PrintChemCondValue,sOut_WSH61)CONCAT(printTreatString[83],sOut_WSH61,sPrntArray[PrintIndex])CONCAT(sPrntArray[PrintIndex],printTreatString[56],sPrntArray[PrintIndex])CONCAT(sPrntArray[PrintIndex],sCRLF,sPrntArray[PrintIndex])[ADD(PrintIndex,1,PrintIndex) ,CLR(PrintChemCondValue) ];
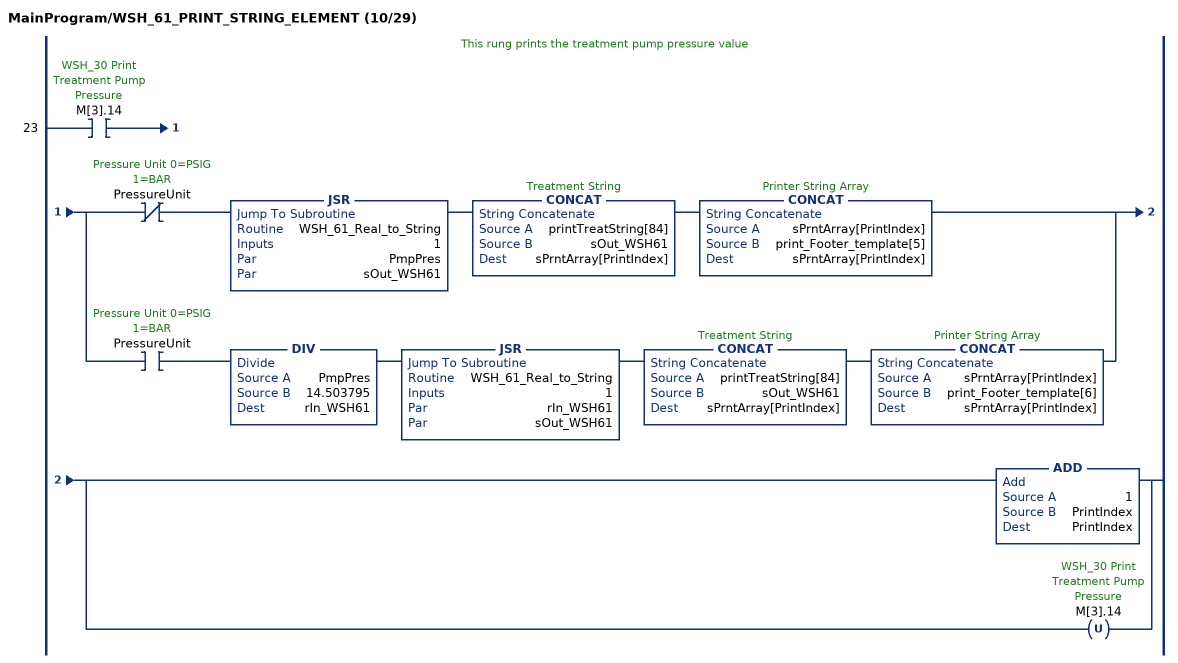
   // This rung prints the treatment pump pressure value
   23: XIC(M[3].14)[XIO(PressureUnit) JSR(WSH_61_Real_to_String,1,PmpPres,sOut_WSH61) CONCAT(printTreatString[84],sOut_WSH61,sPrntArray[PrintIndex]) CONCAT(sPrntArray[PrintIndex],print_Footer_template[5],sPrntArray[PrintIndex]) ,XIC(PressureUnit) DIV(PmpPres,14.503795,rIn_WSH61) JSR(WSH_61_Real_to_String,1,rIn_WSH61,sOut_WSH61) CONCAT(printTreatString[84],sOut_WSH61,sPrntArray[PrintIndex]) CONCAT(sPrntArray[PrintIndex],print_Footer_template[6],sPrntArray[PrintIndex]) ][ADD(1,PrintIndex,PrintIndex) ,OTU(M[3].14) ];
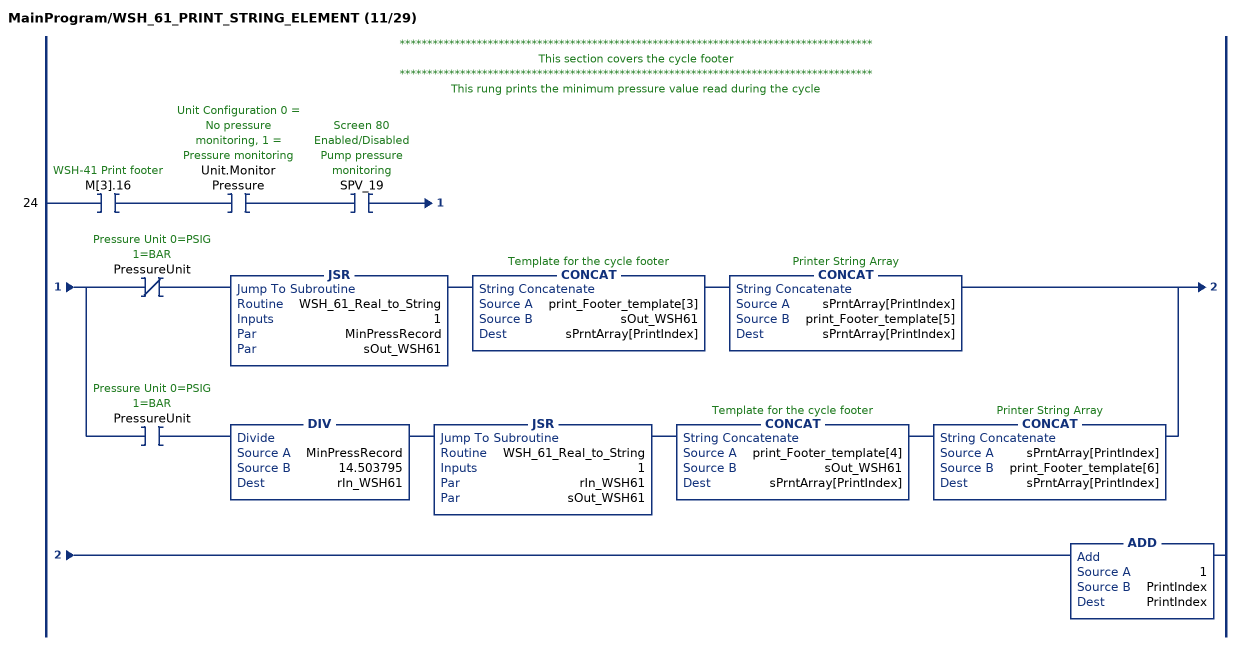
   // **************************************************************************************
   // This section covers the cycle footer
   // **************************************************************************************
   // This rung prints the minimum pressure value read during the cycle
   24: XIC(M[3].16)XIC(Unit.MonitorPressure)XIC(SPV_19)[XIO(PressureUnit) JSR(WSH_61_Real_to_String,1,MinPressRecord,sOut_WSH61) CONCAT(print_Footer_template[3],sOut_WSH61,sPrntArray[PrintIndex]) CONCAT(sPrntArray[PrintIndex],print_Footer_template[5],sPrntArray[PrintIndex]) ,XIC(PressureUnit) DIV(MinPressRecord,14.503795,rIn_WSH61) JSR(WSH_61_Real_to_String,1,rIn_WSH61,sOut_WSH61) CONCAT(print_Footer_template[4],sOut_WSH61,sPrntArray[PrintIndex]) CONCAT(sPrntArray[PrintIndex],print_Footer_template[6],sPrntArray[PrintIndex]) ]ADD(1,PrintIndex,PrintIndex);
